(* PLC project PR_MultiPosShuttle_Soft2.0_Workflow_9b3f4d_PLC, SiemensToBackhoff Siemens TIA Portal to Beckhoff TwinCAT PLCopen Converter 2.0 *)
(* stored: creationDateTime 2026-09-28T09:51:52.682995, modificationDateTime 2026-09-28T09:51:52.682995 *)

FUNCTION_BLOCK PR_MultiPosShuttle_Soft2.0_Workflow_9b3f4d
VAR_INPUT
	iAutoRunning : BOOL;
	iFaultReset : BOOL;
	iGantry2Safe : BOOL;
	iGantry_2Safe : BOOL;
	iHIPOTTesSafe : BOOL;
	iHIPOTTestOver : BOOL;
	iHipotTestInProgress : BOOL;
	iHipotTestSafe : BOOL;
	iInfeedGantrySafe : BOOL;
	iNoRecoveryActive : BOOL;
	iOTS_Frm_Gantry : BOOL;
	iPartPresent : BOOL;
	iPartPrsent : BOOL;
	iPickInProgress : BOOL;
	iPlaceInProgress : BOOL;
	iRTR_Frm_Gantry2 : BOOL;
	iReset_fault : BOOL;
	iShuttleAtGantry2Pos : BOOL;
	iShuttleAtGantry_2Pos : BOOL;
	iShuttleAtHIPOTPos : BOOL;
	iShuttleAtHIPOTTestPos : BOOL;
	iShuttleAtPartLoadPos : BOOL;
	iSstMode : BOOL;
	iSstPB : BOOL;
END_VAR
VAR_OUTPUT
	qError : ARRAY[0..10] OF BOOL;
	qMessage : ARRAY[0..10] OF BOOL;
	qRTR_To_InfeedGantry : BOOL;
	qShuttleGantry_2PosCmd : BOOL;
	qShuttleHIPOTTestPosCmd : BOOL;
	qShuttleReceivePosCmd : BOOL;
END_VAR
VAR
	c10_ChkRecoveryCondition_T1 : BOOL;
	c10_ChkRecoveryCondition_T2 : BOOL;
	c10_ChkRecoveryCondition_T3 : BOOL;
	c10_ChkRecoveryCondition_T4 : BOOL;
	c10_ChkRecoveryCondition_T5 : BOOL;
	c150_ChkOperationStatus_T1 : BOOL;
	c150_ChkOperationStatus_T2 : BOOL;
	c30_ChkPartPresent_T1 : BOOL;
	c30_ChkPartPresent_T2 : BOOL;
	StateNo : INT;
	s100_WtHipotTestOver : BOOL;
	s100_WtHipotTestOver_T1 : BOOL;
	s10_ChkRecoveryCondition : BOOL;
	s10_ChkRecoveryCondition_T1 : BOOL;
	s10_ChkRecoveryCondition_T2 : BOOL;
	s10_ChkRecoveryCondition_T3 : BOOL;
	s10_ChkRecoveryCondition_T4 : BOOL;
	s10_ChkRecoveryCondition_T5 : BOOL;
	s110_WtGantry2AtSafePos : BOOL;
	s110_WtGantry2AtSafePos_T1 : BOOL;
	s120_WtShuttleAtGantry2Pos : BOOL;
	s120_WtShuttleAtGantry2Pos_T1 : BOOL;
	s130_WtRTRFrmGantry2 : BOOL;
	s130_WtRTRFrmGantry2_T1 : BOOL;
	s140_WtPartAbsentGantry2Safe : BOOL;
	s140_WtPartAbsentGantry2Safe_T1 : BOOL;
	s150_ChkOperationStatus : BOOL;
	s150_ChkOperationStatus_T1 : BOOL;
	s150_ChkOperationStatus_T2 : BOOL;
	s1_WtResetRelease : BOOL;
	s1_WtResetRelease_T1 : BOOL;
	s20_WtFaultResetAbnormalCond : BOOL;
	s20_WtFaultResetAbnormalCond_T1 : BOOL;
	s30_ChkPartPresent : BOOL;
	s30_ChkPartPresent_T1 : BOOL;
	s30_ChkPartPresent_T2 : BOOL;
	s40_WtAllSysSafe : BOOL;
	s40_WtAllSysSafe_T1 : BOOL;
	s50_WtShuttleAtPartRcvPos : BOOL;
	s50_WtShuttleAtPartRcvPos_T1 : BOOL;
	s60_WtOTSFrmInfeedGantry : BOOL;
	s60_WtOTSFrmInfeedGantry_T1 : BOOL;
	s70_WtPartPlacedGantrySafe : BOOL;
	s70_WtPartPlacedGantrySafe_T1 : BOOL;
	s80_WtHIPOTTestStnSafe : BOOL;
	s80_WtHIPOTTestStnSafe_T1 : BOOL;
	s90_WtShuttleAtHIPOTTestStn : BOOL;
	s90_WtShuttleAtHIPOTTestStn_T1 : BOOL;
	sHIPOTOprnOver : BOOL;
	sSst : BOOL;
	sSstPulse : BOOL;
	sSstRise : R_TRIG;
	sStWtResetRel : BOOL;
	sStWtResetRel_T1 : BOOL;
END_VAR
VAR_TEMP
	tOne : BOOL;
END_VAR
  VAR  (* added by the conversion: wires and edge detectors of the diagram *)
    _w24 : BOOL;
    _w26 : BOOL;
    _w39 : BOOL;
    _w41 : BOOL;
    _w42 : BOOL;
    _w96 : BOOL;
    _w97 : BOOL;
    _w99 : BOOL;
    _w100 : BOOL;
    _w101 : BOOL;
    _w102 : BOOL;
    _w103 : BOOL;
    _w104 : BOOL;
    _w117 : BOOL;
    _w119 : BOOL;
    _w120 : BOOL;
    _w148 : BOOL;
    _w151 : BOOL;
    _w152 : BOOL;
    _w153 : BOOL;
    _w168 : BOOL;
    _w170 : BOOL;
    _w171 : BOOL;
    _w184 : BOOL;
    _w186 : BOOL;
    _w187 : BOOL;
    _w204 : BOOL;
    _w206 : BOOL;
    _w207 : BOOL;
    _w225 : BOOL;
    _w228 : BOOL;
    _w229 : BOOL;
    _w247 : BOOL;
    _w250 : BOOL;
    _w251 : BOOL;
    _w264 : BOOL;
    _w266 : BOOL;
    _w267 : BOOL;
    _w285 : BOOL;
    _w288 : BOOL;
    _w289 : BOOL;
    _w306 : BOOL;
    _w309 : BOOL;
    _w310 : BOOL;
    _w327 : BOOL;
    _w329 : BOOL;
    _w330 : BOOL;
    _w347 : BOOL;
    _w349 : BOOL;
    _w350 : BOOL;
    _w364 : BOOL;
    _w367 : BOOL;
    _w368 : BOOL;
    _w397 : BOOL;
    _w399 : BOOL;
    _w400 : BOOL;
    _w401 : BOOL;
  END_VAR

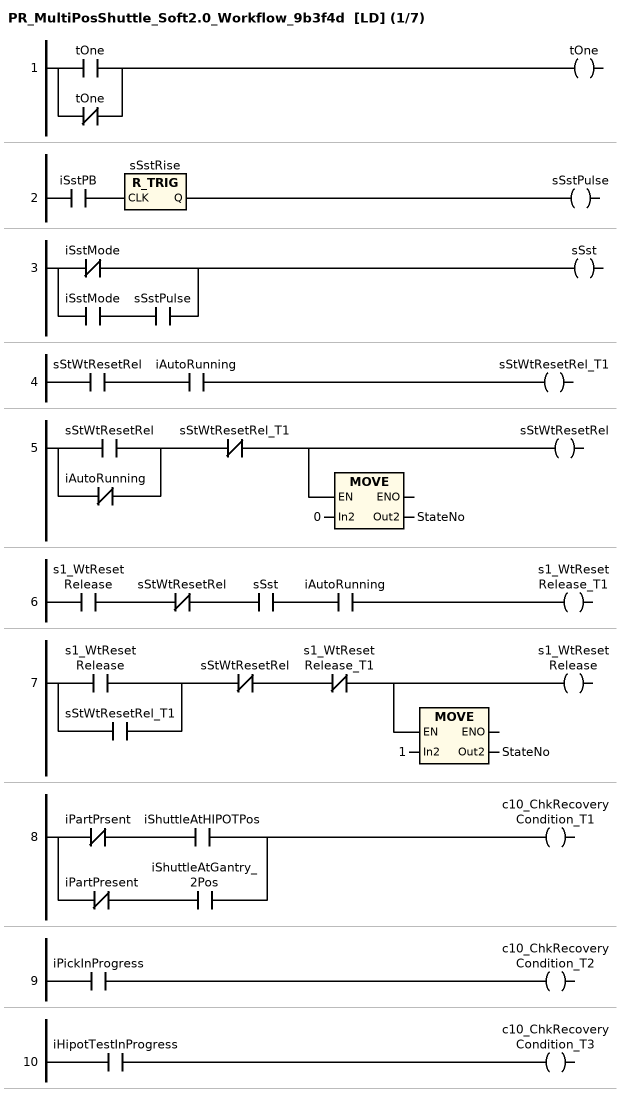
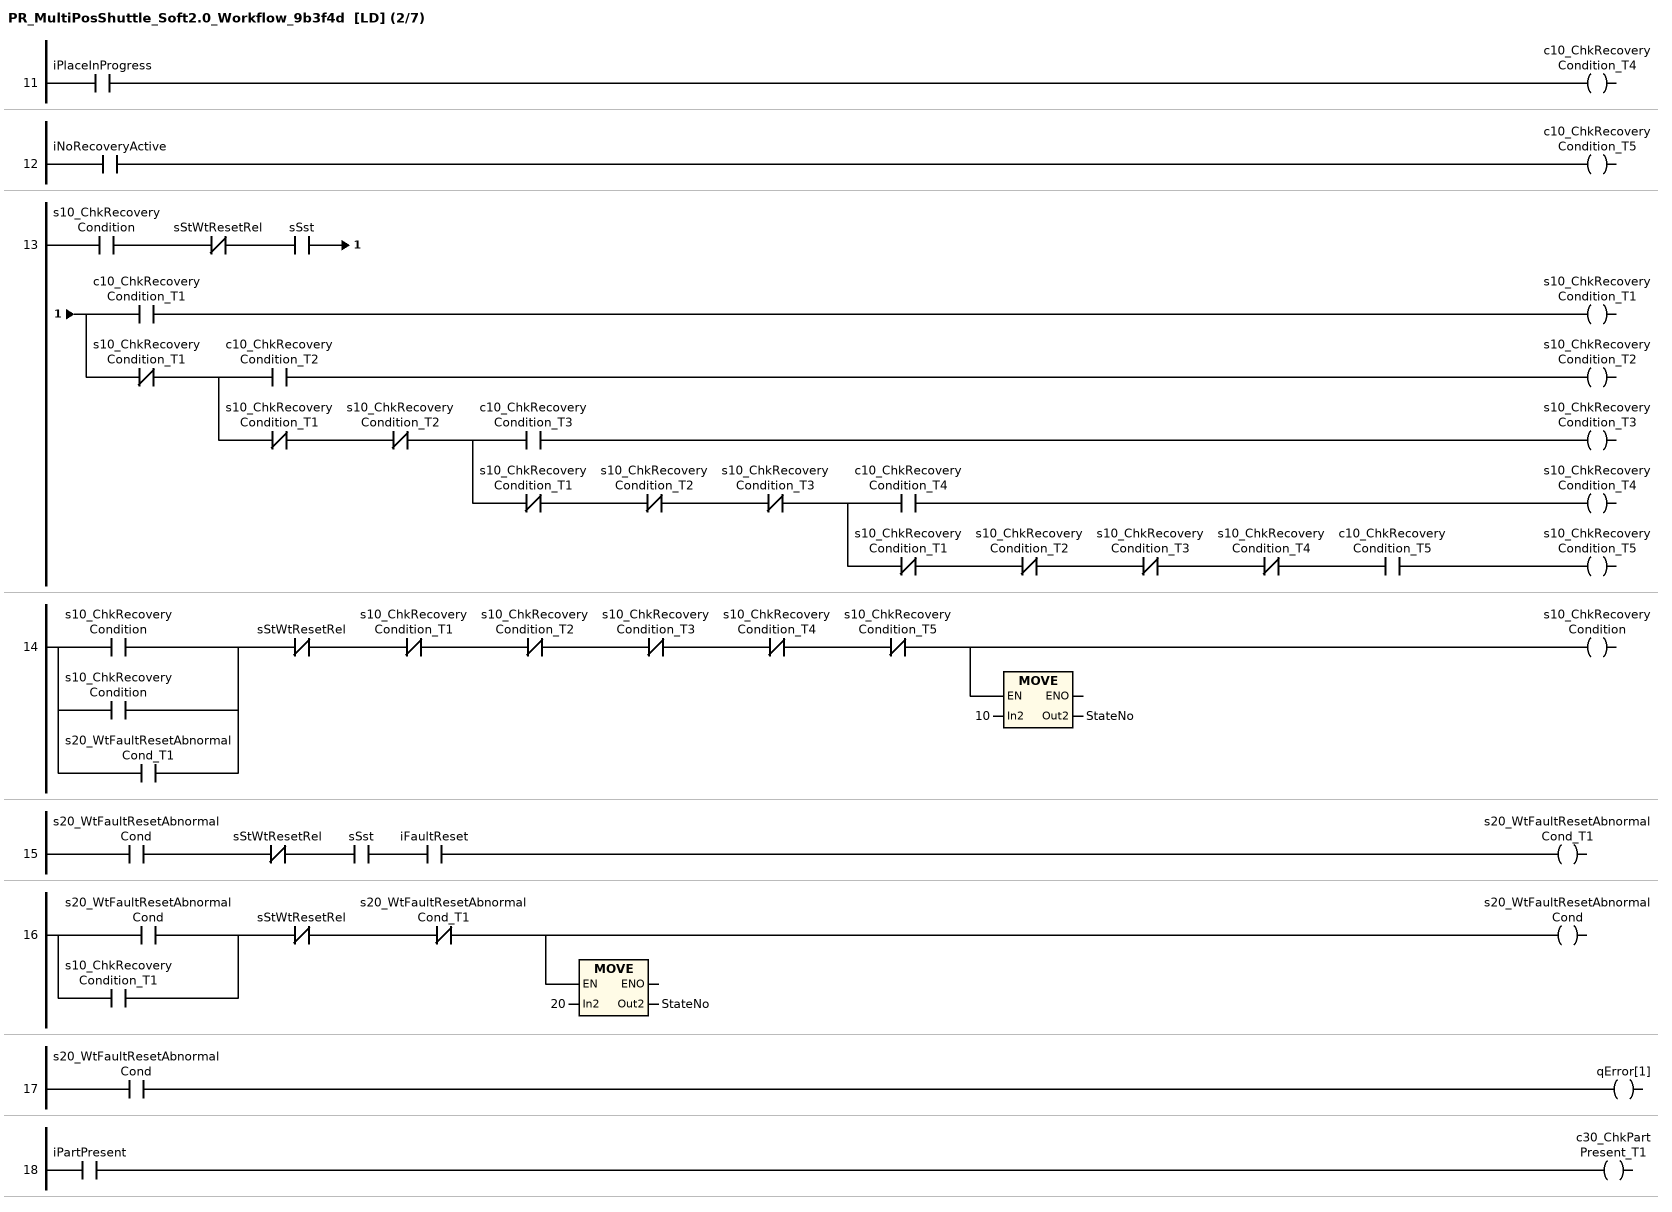
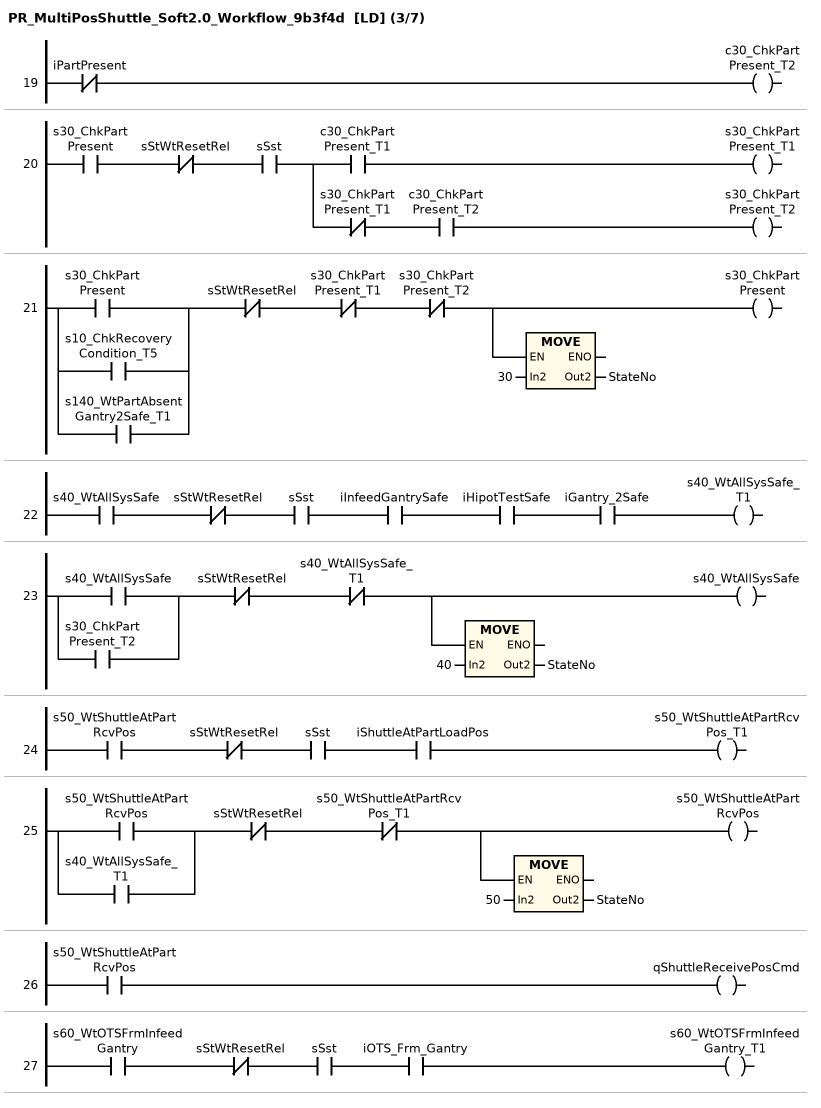
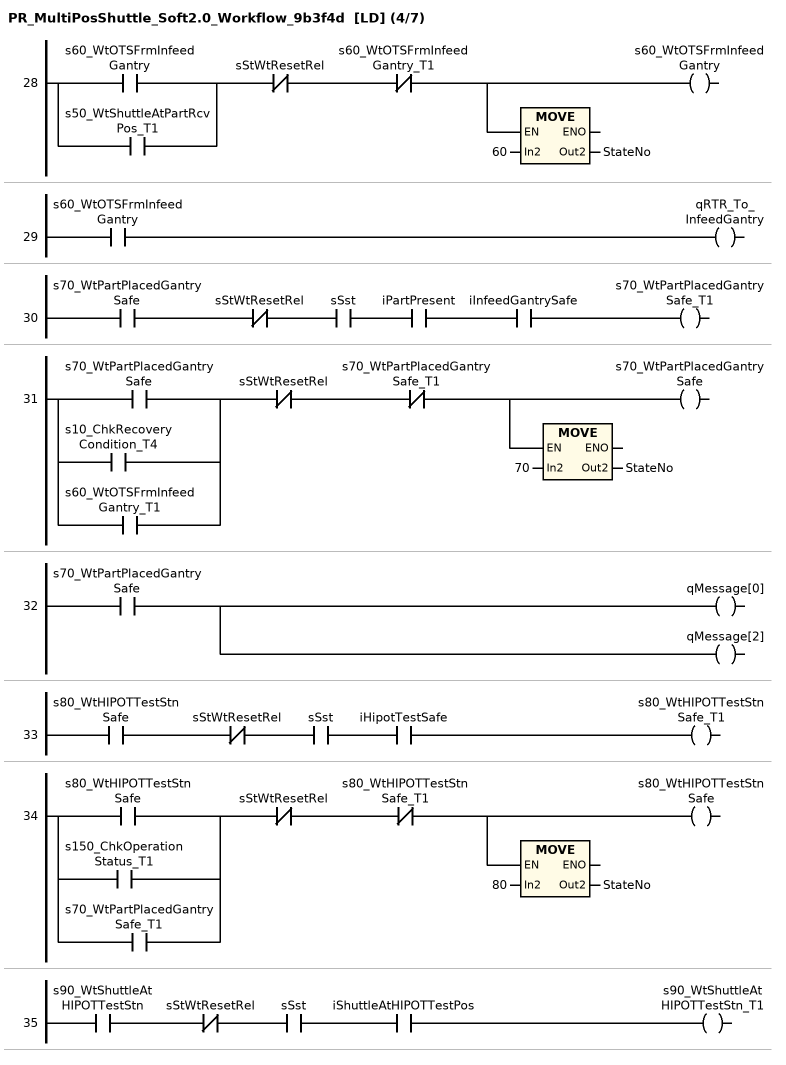
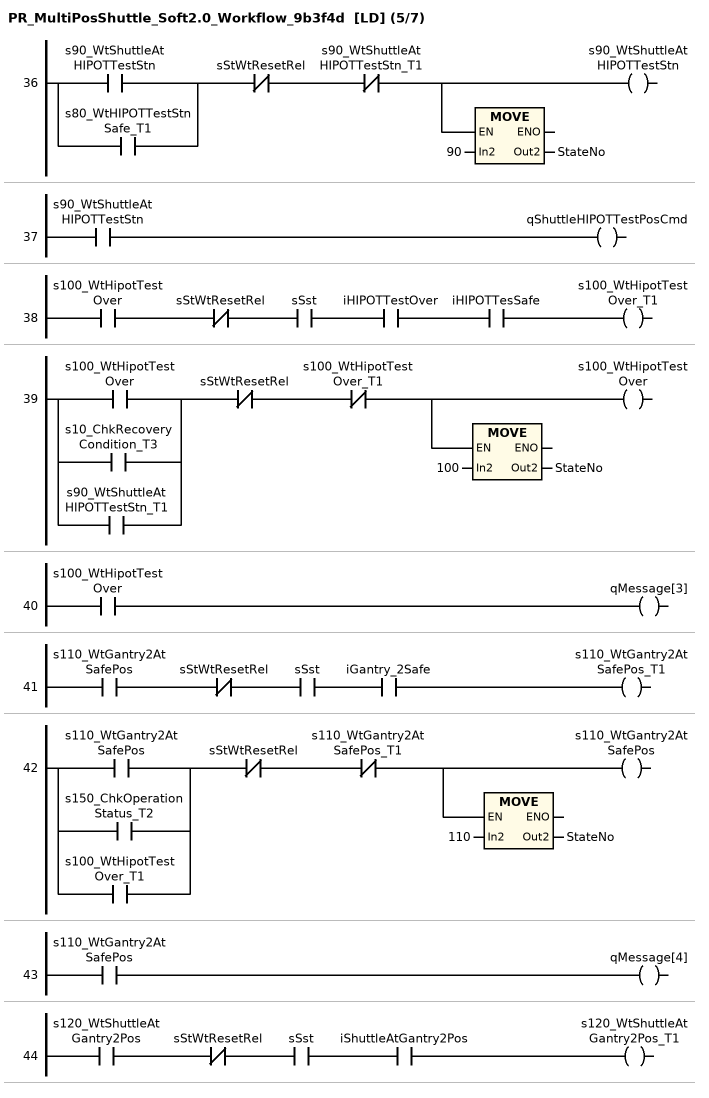
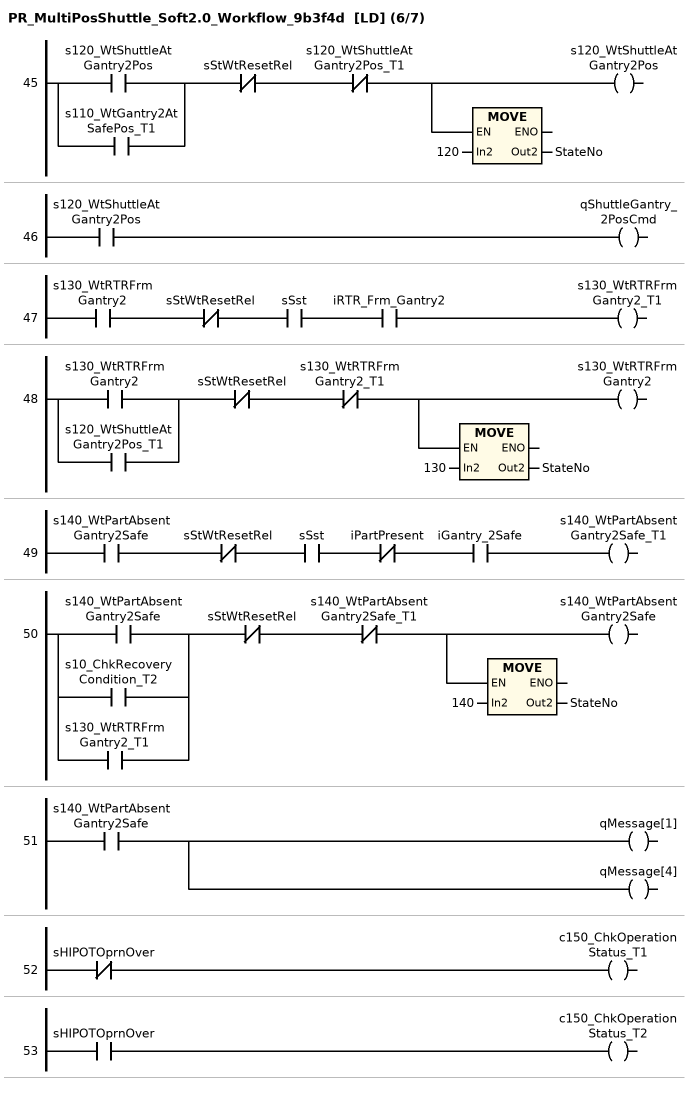
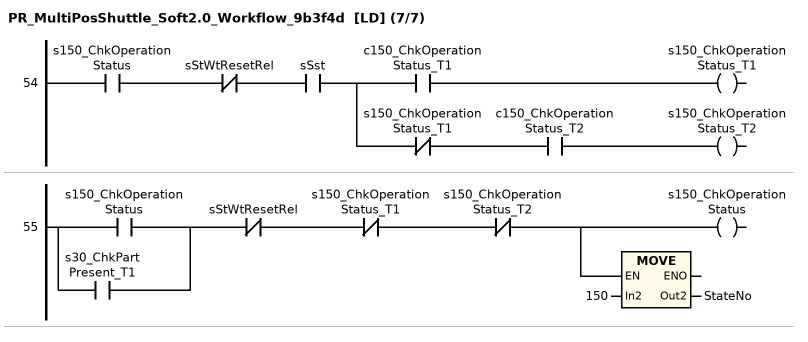
(* LD diagram, written out as Structured Text *)
(* Network 1 *)

tOne := tOne OR NOT tOne;
(* Create Single Step Pulse bit *)

sSstRise(CLK := iSstPB);
sSstPulse := sSstRise.Q;
(* Create Single Step bit *)

sSst := iSstMode AND sSstPulse OR NOT iSstMode;
(* Transition for STATE Num:0 Reset Released *)

sStWtResetRel_T1 := sStWtResetRel AND iAutoRunning;
(* STATE Num:0 Reset Released *)

_w24 := sStWtResetRel;
_w26 := (_w24 OR NOT iAutoRunning) AND NOT sStWtResetRel_T1;
sStWtResetRel := _w26;
IF _w26 THEN StateNo := 0; END_IF;
(* Transition for STATE Num:1 Wait For Reset Release *)

s1_WtResetRelease_T1 := s1_WtResetRelease AND NOT sStWtResetRel AND sSst AND iAutoRunning;
(* STATE Num:1 Wait For Reset Release *)

_w39 := s1_WtResetRelease;
_w41 := (_w39 OR sStWtResetRel_T1) AND NOT sStWtResetRel;
_w42 := _w41 AND NOT s1_WtResetRelease_T1;
s1_WtResetRelease := _w42;
IF _w42 THEN StateNo := 1; END_IF;
(* Condition1 for STATE Num:10 Check Recovery Condition *)

c10_ChkRecoveryCondition_T1 := NOT iPartPrsent AND iShuttleAtHIPOTPos OR NOT iPartPresent AND iShuttleAtGantry_2Pos;
(* Condition2 for STATE Num:10 Check Recovery Condition *)

c10_ChkRecoveryCondition_T2 := iPickInProgress;
(* Condition3 for STATE Num:10 Check Recovery Condition *)

c10_ChkRecoveryCondition_T3 := iHipotTestInProgress;
(* Condition4 for STATE Num:10 Check Recovery Condition *)

c10_ChkRecoveryCondition_T4 := iPlaceInProgress;
(* Condition5 for STATE Num:10 Check Recovery Condition *)

c10_ChkRecoveryCondition_T5 := iNoRecoveryActive;
(* Transition for STATE Num:10 Check Recovery Condition *)

s10_ChkRecoveryCondition_T1 := s10_ChkRecoveryCondition AND NOT sStWtResetRel AND sSst AND c10_ChkRecoveryCondition_T1;
s10_ChkRecoveryCondition_T2 := s10_ChkRecoveryCondition AND NOT sStWtResetRel AND sSst AND NOT s10_ChkRecoveryCondition_T1 AND c10_ChkRecoveryCondition_T2;
s10_ChkRecoveryCondition_T3 := s10_ChkRecoveryCondition AND NOT sStWtResetRel AND sSst AND NOT s10_ChkRecoveryCondition_T1 AND NOT s10_ChkRecoveryCondition_T1 AND NOT s10_ChkRecoveryCondition_T2 AND c10_ChkRecoveryCondition_T3;
s10_ChkRecoveryCondition_T4 := s10_ChkRecoveryCondition AND NOT sStWtResetRel AND sSst AND NOT s10_ChkRecoveryCondition_T1 AND NOT s10_ChkRecoveryCondition_T1 AND NOT s10_ChkRecoveryCondition_T2 AND NOT s10_ChkRecoveryCondition_T1 AND NOT s10_ChkRecoveryCondition_T2 AND NOT s10_ChkRecoveryCondition_T3 AND c10_ChkRecoveryCondition_T4;
s10_ChkRecoveryCondition_T5 := s10_ChkRecoveryCondition AND NOT sStWtResetRel AND sSst AND NOT s10_ChkRecoveryCondition_T1 AND NOT s10_ChkRecoveryCondition_T1 AND NOT s10_ChkRecoveryCondition_T2 AND NOT s10_ChkRecoveryCondition_T1 AND NOT s10_ChkRecoveryCondition_T2 AND NOT s10_ChkRecoveryCondition_T3 AND NOT s10_ChkRecoveryCondition_T1 AND NOT s10_ChkRecoveryCondition_T2 AND NOT s10_ChkRecoveryCondition_T3 AND NOT s10_ChkRecoveryCondition_T4 AND c10_ChkRecoveryCondition_T5;
(* STATE Num:10 Check Recovery Condition *)

_w96 := s10_ChkRecoveryCondition;
_w97 := s10_ChkRecoveryCondition;
_w99 := (_w96 OR _w97 OR s20_WtFaultResetAbnormalCond_T1) AND NOT sStWtResetRel;
_w100 := _w99 AND NOT s10_ChkRecoveryCondition_T1;
_w101 := _w100 AND NOT s10_ChkRecoveryCondition_T2;
_w102 := _w101 AND NOT s10_ChkRecoveryCondition_T3;
_w103 := _w102 AND NOT s10_ChkRecoveryCondition_T4;
_w104 := _w103 AND NOT s10_ChkRecoveryCondition_T5;
s10_ChkRecoveryCondition := _w104;
IF _w104 THEN StateNo := 10; END_IF;
(* Transition for STATE Num:20 Wait for Fault Reset_AbnormalCond *)

s20_WtFaultResetAbnormalCond_T1 := s20_WtFaultResetAbnormalCond AND NOT sStWtResetRel AND sSst AND iFaultReset;
(* STATE Num:20 Wait for Fault Reset_AbnormalCond *)

_w117 := s20_WtFaultResetAbnormalCond;
_w119 := (_w117 OR s10_ChkRecoveryCondition_T1) AND NOT sStWtResetRel;
_w120 := _w119 AND NOT s20_WtFaultResetAbnormalCond_T1;
s20_WtFaultResetAbnormalCond := _w120;
IF _w120 THEN StateNo := 20; END_IF;
(* Actions for STATE Num:20 Wait for Fault Reset_AbnormalCond *)

qError[1] := s20_WtFaultResetAbnormalCond;
(* Condition1 for STATE Num:30 Check Part Present *)

c30_ChkPartPresent_T1 := iPartPresent;
(* Condition2 for STATE Num:30 Check Part Present *)

c30_ChkPartPresent_T2 := NOT iPartPresent;
(* Transition for STATE Num:30 Check Part Present *)

s30_ChkPartPresent_T1 := s30_ChkPartPresent AND NOT sStWtResetRel AND sSst AND c30_ChkPartPresent_T1;
s30_ChkPartPresent_T2 := s30_ChkPartPresent AND NOT sStWtResetRel AND sSst AND NOT s30_ChkPartPresent_T1 AND c30_ChkPartPresent_T2;
(* STATE Num:30 Check Part Present *)

_w148 := s30_ChkPartPresent;
_w151 := (_w148 OR s10_ChkRecoveryCondition_T5 OR s140_WtPartAbsentGantry2Safe_T1) AND NOT sStWtResetRel;
_w152 := _w151 AND NOT s30_ChkPartPresent_T1;
_w153 := _w152 AND NOT s30_ChkPartPresent_T2;
s30_ChkPartPresent := _w153;
IF _w153 THEN StateNo := 30; END_IF;
(* Transition for STATE Num:40 Wait All System Safe for Shuttle Motion *)

s40_WtAllSysSafe_T1 := s40_WtAllSysSafe AND NOT sStWtResetRel AND sSst AND iInfeedGantrySafe AND iHipotTestSafe AND iGantry_2Safe;
(* STATE Num:40 Wait All System Safe for Shuttle Motion *)

_w168 := s40_WtAllSysSafe;
_w170 := (_w168 OR s30_ChkPartPresent_T2) AND NOT sStWtResetRel;
_w171 := _w170 AND NOT s40_WtAllSysSafe_T1;
s40_WtAllSysSafe := _w171;
IF _w171 THEN StateNo := 40; END_IF;
(* Transition for STATE Num:50 Wait for Shuttle At Part Receive Pos *)

s50_WtShuttleAtPartRcvPos_T1 := s50_WtShuttleAtPartRcvPos AND NOT sStWtResetRel AND sSst AND iShuttleAtPartLoadPos;
(* STATE Num:50 Wait for Shuttle At Part Receive Pos *)

_w184 := s50_WtShuttleAtPartRcvPos;
_w186 := (_w184 OR s40_WtAllSysSafe_T1) AND NOT sStWtResetRel;
_w187 := _w186 AND NOT s50_WtShuttleAtPartRcvPos_T1;
s50_WtShuttleAtPartRcvPos := _w187;
IF _w187 THEN StateNo := 50; END_IF;
(* Actions for STATE Num:50 Wait for Shuttle At Part Receive Pos *)

qShuttleReceivePosCmd := s50_WtShuttleAtPartRcvPos;
(* Transition for STATE Num:60 Wait for OTS From Infeed Gantry *)

s60_WtOTSFrmInfeedGantry_T1 := s60_WtOTSFrmInfeedGantry AND NOT sStWtResetRel AND sSst AND iOTS_Frm_Gantry;
(* STATE Num:60 Wait for OTS From Infeed Gantry *)

_w204 := s60_WtOTSFrmInfeedGantry;
_w206 := (_w204 OR s50_WtShuttleAtPartRcvPos_T1) AND NOT sStWtResetRel;
_w207 := _w206 AND NOT s60_WtOTSFrmInfeedGantry_T1;
s60_WtOTSFrmInfeedGantry := _w207;
IF _w207 THEN StateNo := 60; END_IF;
(* Actions for STATE Num:60 Wait for OTS From Infeed Gantry *)

qRTR_To_InfeedGantry := s60_WtOTSFrmInfeedGantry;
(* Transition for STATE Num:70 Wait for part Placed By Gantry and Gantry Safe *)

s70_WtPartPlacedGantrySafe_T1 := s70_WtPartPlacedGantrySafe AND NOT sStWtResetRel AND sSst AND iPartPresent AND iInfeedGantrySafe;
(* STATE Num:70 Wait for part Placed By Gantry and Gantry Safe *)

_w225 := s70_WtPartPlacedGantrySafe;
_w228 := (_w225 OR s10_ChkRecoveryCondition_T4 OR s60_WtOTSFrmInfeedGantry_T1) AND NOT sStWtResetRel;
_w229 := _w228 AND NOT s70_WtPartPlacedGantrySafe_T1;
s70_WtPartPlacedGantrySafe := _w229;
IF _w229 THEN StateNo := 70; END_IF;
(* Actions for STATE Num:70 Wait for part Placed By Gantry and Gantry Safe *)

qMessage[0] := s70_WtPartPlacedGantrySafe;
qMessage[2] := s70_WtPartPlacedGantrySafe;
(* Transition for STATE Num:80 Wait for HIPOT Test Station Safe *)

s80_WtHIPOTTestStnSafe_T1 := s80_WtHIPOTTestStnSafe AND NOT sStWtResetRel AND sSst AND iHipotTestSafe;
(* STATE Num:80 Wait for HIPOT Test Station Safe *)

_w247 := s80_WtHIPOTTestStnSafe;
_w250 := (_w247 OR s150_ChkOperationStatus_T1 OR s70_WtPartPlacedGantrySafe_T1) AND NOT sStWtResetRel;
_w251 := _w250 AND NOT s80_WtHIPOTTestStnSafe_T1;
s80_WtHIPOTTestStnSafe := _w251;
IF _w251 THEN StateNo := 80; END_IF;
(* Transition for STATE Num:90 Wait for Shuttle at HIPOT Test Station *)

s90_WtShuttleAtHIPOTTestStn_T1 := s90_WtShuttleAtHIPOTTestStn AND NOT sStWtResetRel AND sSst AND iShuttleAtHIPOTTestPos;
(* STATE Num:90 Wait for Shuttle at HIPOT Test Station *)

_w264 := s90_WtShuttleAtHIPOTTestStn;
_w266 := (_w264 OR s80_WtHIPOTTestStnSafe_T1) AND NOT sStWtResetRel;
_w267 := _w266 AND NOT s90_WtShuttleAtHIPOTTestStn_T1;
s90_WtShuttleAtHIPOTTestStn := _w267;
IF _w267 THEN StateNo := 90; END_IF;
(* Actions for STATE Num:90 Wait for Shuttle at HIPOT Test Station *)

qShuttleHIPOTTestPosCmd := s90_WtShuttleAtHIPOTTestStn;
(* Transition for STATE Num:100 Wait for Hipot Test Over *)

s100_WtHipotTestOver_T1 := s100_WtHipotTestOver AND NOT sStWtResetRel AND sSst AND iHIPOTTestOver AND iHIPOTTesSafe;
(* STATE Num:100 Wait for Hipot Test Over *)

_w285 := s100_WtHipotTestOver;
_w288 := (_w285 OR s10_ChkRecoveryCondition_T3 OR s90_WtShuttleAtHIPOTTestStn_T1) AND NOT sStWtResetRel;
_w289 := _w288 AND NOT s100_WtHipotTestOver_T1;
s100_WtHipotTestOver := _w289;
IF _w289 THEN StateNo := 100; END_IF;
(* Actions for STATE Num:100 Wait for Hipot Test Over *)

qMessage[3] := s100_WtHipotTestOver;
(* Transition for STATE Num:110 Wait for Gantry-2 At Safe Position *)

s110_WtGantry2AtSafePos_T1 := s110_WtGantry2AtSafePos AND NOT sStWtResetRel AND sSst AND iGantry_2Safe;
(* STATE Num:110 Wait for Gantry-2 At Safe Position *)

_w306 := s110_WtGantry2AtSafePos;
_w309 := (_w306 OR s150_ChkOperationStatus_T2 OR s100_WtHipotTestOver_T1) AND NOT sStWtResetRel;
_w310 := _w309 AND NOT s110_WtGantry2AtSafePos_T1;
s110_WtGantry2AtSafePos := _w310;
IF _w310 THEN StateNo := 110; END_IF;
(* Actions for STATE Num:110 Wait for Gantry-2 At Safe Position *)

qMessage[4] := s110_WtGantry2AtSafePos;
(* Transition for STATE Num:120 Wait Shuttle at Gantry-2 Position *)

s120_WtShuttleAtGantry2Pos_T1 := s120_WtShuttleAtGantry2Pos AND NOT sStWtResetRel AND sSst AND iShuttleAtGantry2Pos;
(* STATE Num:120 Wait Shuttle at Gantry-2 Position *)

_w327 := s120_WtShuttleAtGantry2Pos;
_w329 := (_w327 OR s110_WtGantry2AtSafePos_T1) AND NOT sStWtResetRel;
_w330 := _w329 AND NOT s120_WtShuttleAtGantry2Pos_T1;
s120_WtShuttleAtGantry2Pos := _w330;
IF _w330 THEN StateNo := 120; END_IF;
(* Actions for STATE Num:120 Wait Shuttle at Gantry-2 Position *)

qShuttleGantry_2PosCmd := s120_WtShuttleAtGantry2Pos;
(* Transition for STATE Num:130 Wait RTR From Gantry-2 *)

s130_WtRTRFrmGantry2_T1 := s130_WtRTRFrmGantry2 AND NOT sStWtResetRel AND sSst AND iRTR_Frm_Gantry2;
(* STATE Num:130 Wait RTR From Gantry-2 *)

_w347 := s130_WtRTRFrmGantry2;
_w349 := (_w347 OR s120_WtShuttleAtGantry2Pos_T1) AND NOT sStWtResetRel;
_w350 := _w349 AND NOT s130_WtRTRFrmGantry2_T1;
s130_WtRTRFrmGantry2 := _w350;
IF _w350 THEN StateNo := 130; END_IF;
(* Transition for STATE Num:140 Wait for Part Absent and Gantry-2 safe *)

s140_WtPartAbsentGantry2Safe_T1 := s140_WtPartAbsentGantry2Safe AND NOT sStWtResetRel AND sSst AND NOT iPartPresent AND iGantry_2Safe;
(* STATE Num:140 Wait for Part Absent and Gantry-2 safe *)

_w364 := s140_WtPartAbsentGantry2Safe;
_w367 := (_w364 OR s10_ChkRecoveryCondition_T2 OR s130_WtRTRFrmGantry2_T1) AND NOT sStWtResetRel;
_w368 := _w367 AND NOT s140_WtPartAbsentGantry2Safe_T1;
s140_WtPartAbsentGantry2Safe := _w368;
IF _w368 THEN StateNo := 140; END_IF;
(* Actions for STATE Num:140 Wait for Part Absent and Gantry-2 safe *)

qMessage[1] := s140_WtPartAbsentGantry2Safe;
qMessage[4] := s140_WtPartAbsentGantry2Safe;
(* Condition1 for STATE Num:150 Check Operation Status *)

c150_ChkOperationStatus_T1 := NOT sHIPOTOprnOver;
(* Condition2 for STATE Num:150 Check Operation Status *)

c150_ChkOperationStatus_T2 := sHIPOTOprnOver;
(* Transition for STATE Num:150 Check Operation Status *)

s150_ChkOperationStatus_T1 := s150_ChkOperationStatus AND NOT sStWtResetRel AND sSst AND c150_ChkOperationStatus_T1;
s150_ChkOperationStatus_T2 := s150_ChkOperationStatus AND NOT sStWtResetRel AND sSst AND NOT s150_ChkOperationStatus_T1 AND c150_ChkOperationStatus_T2;
(* STATE Num:150 Check Operation Status *)

_w397 := s150_ChkOperationStatus;
_w399 := (_w397 OR s30_ChkPartPresent_T1) AND NOT sStWtResetRel;
_w400 := _w399 AND NOT s150_ChkOperationStatus_T1;
_w401 := _w400 AND NOT s150_ChkOperationStatus_T2;
s150_ChkOperationStatus := _w401;
IF _w401 THEN StateNo := 150; END_IF;
END_FUNCTION_BLOCK
